SUBAPPLICATION AUF_AB_Button_BG (* Manuell Auf/Ab mit 2 Buttons, nur Anzeige und AX-Ausgaenge (ohne eigene Ventilausgaenge) *)
  (* Standard: 61499-2; Description: Copyright (c) 2026 Meisterschulen am Ostbahnhof This program and the accompanying materials are made available under the terms of the Eclipse Public License 2.0 which is available at https://www.eclipse.org/legal/epl-2.0/ SPDX-License-Identifier: EPL-2.0 *)
  (* Version 1.0, 2026-10-31, Franz Höpfinger, Meisterschulen am Ostbahnhof, Aus Getreidehacke func/Manual/ManFunc_AUF_AB0 in MyLib::sys verschoben und umbenannt, INIT/INITO/QI/QO ergaenzt. *)
  PACKAGE MyLib::sys;
  IMPORT isobus::UT::Q::const::IDs::ID_NULL;
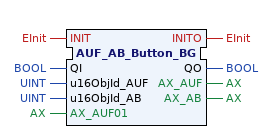
  EVENT_INPUT
    INIT : EInit; (* Initialization Request *)
  END_EVENT
  EVENT_OUTPUT
    INITO : EInit; (* Initialization Confirm *)
  END_EVENT
  VAR_INPUT
    QI : BOOL := TRUE; (* Quality Input - TRUE to enable service *)
    u16ObjId_AUF : UINT := ID_NULL; (* Object ID Button AUF *)
    u16ObjId_AB : UINT := ID_NULL; (* Object ID Button AB *)
  END_VAR
  VAR_OUTPUT
    QO : BOOL; (* Quality Output - TRUE if service executed successfully *)
  END_VAR
  SOCKETS
    AX_AUF01 : adapter::types::unidirectional::AX; (* externer Eingang AUF *)
  END_SOCKETS
  PLUGS
    AX_AUF : adapter::types::unidirectional::AX; (* AUF aktiv *)
    AX_AB : adapter::types::unidirectional::AX; (* AB aktiv *)
  END_PLUGS
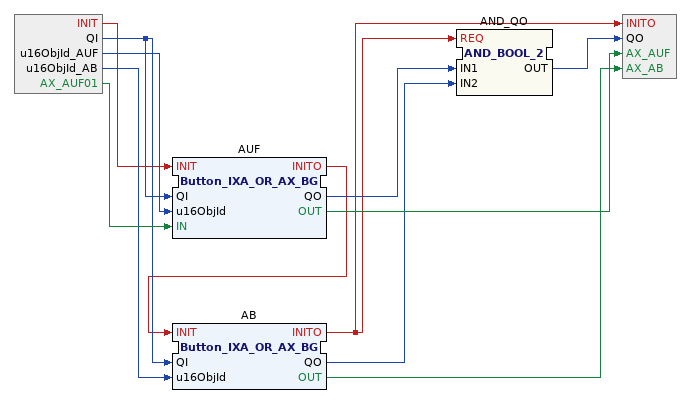
  FBS
    AND_QO : iec61131::booleanOperators::AND_BOOL_2;
  END_FBS
  SUBAPPS
    AUF : MyLib::sys::Button_IXA_OR_AX_BG;
    AB : MyLib::sys::Button_IXA_OR_AX_BG;
  END_SUBAPPS
  EVENT_CONNECTIONS
    INIT TO AUF.INIT;
    AUF.INITO TO AB.INIT;
    AB.INITO TO INITO;
    AB.INITO TO AND_QO.REQ;
  END_CONNECTIONS
  DATA_CONNECTIONS
    QI TO AUF.QI;
    QI TO AB.QI;
    u16ObjId_AUF TO AUF.u16ObjId;
    u16ObjId_AB TO AB.u16ObjId;
    AUF.QO TO AND_QO.IN1;
    AB.QO TO AND_QO.IN2;
    AND_QO.OUT TO QO;
  END_CONNECTIONS
  ADAPTER_CONNECTIONS
    AX_AUF01 TO AUF.IN;
    AUF.OUT TO AX_AUF;
    AB.OUT TO AX_AB;
  END_CONNECTIONS
END_SUBAPPLICATION
